TYPE ST_PolarIIChamber_ArmRotateServiceCtrl :
STRUCT
	JogPositive : ST_ServiceCtrl;
	JogNegative : ST_ServiceCtrl;
	IncrementalJog : ST_ServiceCtrl;
	MoveRecipe : ST_ServiceCtrl;
	NegLimitPos : ST_ServiceCtrl;
	PosLimitPos : ST_ServiceCtrl;
	NozzlePortPos : ST_ServiceCtrl;
	Noz1CenterPos : ST_ServiceCtrl;
	Noz2CenterPos : ST_ServiceCtrl;
	Noz3CenterPos : ST_ServiceCtrl;
END_STRUCT
END_TYPE

(* stored: Version 1.1.0.1, ProductVersion 3.1.4026.18
   DUT ST_PolarIIChamber_ArmRotateServiceCtrl: Id {14000000-0000-0000-0000-000000000025} *)
